(* CODESYS project tcprocess.library
   Company: TcNexa
   DefaultNamespace: TcNexa_Components_TcProcess
   Version: 1.0.0.0
   Placeholder: TcProcess
   Author: ATI Software Engineering
   Description: This library serves as a valuable resource for managing reusable components within your automation projects
   Title: TcProcess

Project tree, tasks and I/O mapping:
  libraries: Tc2_Standard, * (Beckhoff Automation GmbH); Tc2_System, * (Beckhoff Automation GmbH); Tc3_Module, * (Beckhoff Automation GmbH)
  Method Reponse/
    function block FB_MethodResponse [ST]: _clear, busy, description, error, copyFrom, setBusy, setFail, setPass
  Step/
    function block FB_Step [ST]: actual, inc, init, set
  Tests/
    program PRG_TEST [ST]
  Version/
    global variables Global_Version
*)

// Version/Global_Version
{attribute 'TcGenerated'}
{attribute 'no-analysis'}
{attribute 'linkalways'}
// This function has been automatically generated from the project information.
VAR_GLOBAL CONSTANT
	{attribute 'const_non_replaced'}
	stLibVersion_TcProcess : ST_LibVersion := (iMajor := 1, iMinor := 0, iBuild := 0, iRevision := 0, nFlags := 0, sVersion := '1.0.0.0');
END_VAR

// Method Reponse/FB_MethodResponse
FUNCTION_BLOCK FB_MethodResponse
VAR
	_busy			: BOOL;						// Indicates if the method call is in progress
	_error			: BOOL;						// Indicates if the method call failed
	_description	: Tc2_System.T_MaxString;	// Information to show to the user
	
	
	
	
//	_statusMsg		: Tc2_System.T_MaxString;	// Status message from method call
//	_statusId		: UDINT;					// Message ID from method call, for further processing (translation etc.)
//	_errorMsg		: Tc2_System.T_MaxString;	// Error message from method call
//	_errorId		: UDINT;					// Error ID from method call
//	_errorSrc		: STRING;					// Source for the error (Beckhoff, Keyence etc.)
END_VAR

METHOD PROTECTED _clear
VAR_INPUT
END_VAR
_busy:= FALSE;
_error:= FALSE;
_description:= '';
END_METHOD

PROPERTY PUBLIC busy : BOOL
GET
busy:= _busy;
END_GET
END_PROPERTY

PROPERTY PUBLIC description : Tc2_System.T_MaxString
GET
description:= _description;
END_GET
END_PROPERTY

PROPERTY PUBLIC error : BOOL
GET
error:= _error;
END_GET
END_PROPERTY

METHOD PUBLIC copyFrom
VAR_INPUT
	Response		: FB_MethodResponse;
END_VAR
_busy:= Response.busy;
_error:= Response.error;
_description:= Response.description;
END_METHOD

METHOD PUBLIC setBusy
VAR_INPUT
	description	 	: Tc2_System.T_MaxString;
END_VAR
_clear();

_busy:= TRUE;
_description:= description;
END_METHOD

METHOD PUBLIC setFail
VAR_INPUT
	description	 	: Tc2_System.T_MaxString;
END_VAR
_clear();

_error:= TRUE;
_description:= description;
END_METHOD

METHOD PUBLIC setPass
VAR_INPUT
END_VAR
_clear();
END_METHOD

END_FUNCTION_BLOCK

// Step/FB_Step
FUNCTION_BLOCK FB_Step
VAR
	_actual						: INT:= -1;
END_VAR

PROPERTY PUBLIC actual : INT
GET
PUBLIC 
VAR
END_VAR
actual:= _actual;
END_GET
END_PROPERTY

METHOD PUBLIC inc
VAR
END_VAR
_actual:= _actual + 1;
END_METHOD

METHOD PUBLIC init
VAR_INPUT
END_VAR
_actual:= 0;
END_METHOD

METHOD PUBLIC set
VAR_INPUT
	target	: INT;
END_VAR
_actual:= target;
END_METHOD

END_FUNCTION_BLOCK

// Tests/PRG_TEST
PROGRAM PRG_TEST
VAR
END_VAR

END_PROGRAM
